// TIA Portal project "000_empty" (V21)

(* hardware
DEVICE "PLC_1"  S7-1500 station
   slot 0: "Rail_0"  Rack  6ES7 590-1***0-0AA0
   slot 1: "PLC_1"  CPU 1513-1 PN  6ES7 513-1AL02-0AB0  V2.9
      slot 3: "CPU display_1"  6ES7591-1AA00-0AA0
      slot 32768: "PROFINET interface_1"  X1
         slot 32769: "Port_1"  X1 P1
         slot 32770: "Port_2"  X1 P2
      slot 34817: "Virtual CP interface port_1"  Virtual CP interface port  Virtual CP interface port
*)

// ===== PLC "PLC_1"  CPU 1513-1 PN =====

TYPE "UDT_Motor"
   STRUCT
      Running : Bool;   // Motor on
      Speed : Real := 1500.0;   // Speed setpoint
      Count : Int := 7;
   END_STRUCT;
END_TYPE

DATA_BLOCK "DB_Global"   // DB1
{ S7_Optimized_Access := 'TRUE' }
   VAR
      xBool : Bool := TRUE;   // Bool comment
      iInt : Int := 42;
      rReal : Real := 3.5;   // Real comment
      aInt : Array[0..3] of Int;
      sData : Struct
         "a" : Bool;
         "b" : DInt := -5;
      END_STRUCT;
   END_VAR
BEGIN
   aInt[1] := 11;
END_DATA_BLOCK

DATA_BLOCK "FB_Empty_DB"   // DB2
{ S7_Optimized_Access := 'TRUE' }
VERSION : 0.1
// stored: InstanceOfName FB_Empty
"FB_Empty"
BEGIN
END_DATA_BLOCK

DATA_BLOCK "DB_Motor"   // DB4
{ S7_Optimized_Access := 'TRUE' }
   VAR
      motor : "UDT_Motor";
   END_VAR
BEGIN
   motor.Speed := 750.0;
END_DATA_BLOCK

// folder: BlockGroup_1

DATA_BLOCK "DB_InGroup"   // DB3
{ S7_Optimized_Access := 'TRUE' }
   VAR
      wWord : Word := 16#00FF;
   END_VAR
BEGIN
END_DATA_BLOCK

// folder: (top level)

FUNCTION_BLOCK "FB_Empty"   // FB1, SCL
{ S7_Optimized_Access := 'TRUE' }
VERSION : 0.1
BEGIN
END_FUNCTION_BLOCK

FUNCTION_BLOCK "FB_Iface"   // FB2, SCL
{ S7_Optimized_Access := 'TRUE' }
VERSION : 0.1
   VAR_INPUT
      iBool : Bool;   // Input bool
      iInt : Int;   // Input int
      iReal : Real;   // Input real
      iArr : Array[0..3] of Int;   // Input array
      iMotor : "UDT_Motor";   // Input UDT
   END_VAR
   VAR_OUTPUT
      oBool : Bool;   // Output bool
      oInt : Int;   // Output int
   END_VAR
   VAR_IN_OUT
      ioReal : Real;   // InOut real
   END_VAR
   VAR
      stInt : Int := 42;   // Static int
      stBool : Bool;   // Static bool comment
   END_VAR
   VAR_TEMP
      tInt : Int;   // Temp int
   END_VAR
   VAR CONSTANT
      cInt : Int := 7;   // Constant int
   END_VAR
BEGIN
   #tInt := #iInt + #cInt;
           #oInt := #tInt;
           #oBool := #iBool;
           #ioReal := #ioReal + #iReal;
END_FUNCTION_BLOCK

FUNCTION "FC_Iface" : Int   // FC1, SCL
{ S7_Optimized_Access := 'TRUE' }
VERSION : 0.1
   VAR_INPUT
      iBool : Bool;   // Input bool
      iInt : Int;   // Input int
      iReal : Real;   // Input real
      iArr : Array[0..3] of Int;   // Input array
      iMotor : "UDT_Motor";   // Input UDT
   END_VAR
   VAR_OUTPUT
      oBool : Bool;   // Output bool
      oInt : Int;   // Output int
   END_VAR
   VAR_IN_OUT
      ioReal : Real;   // InOut real
   END_VAR
   VAR_TEMP
      tInt : Int;   // Temp int
   END_VAR
   VAR CONSTANT
      cInt : Int := 7;   // Constant int
   END_VAR
BEGIN
   #tInt := #iInt + #cInt;
           #oInt := #tInt;
           #oBool := #iBool;
           #ioReal := #ioReal + #iReal;
           #FC_Iface := #tInt;
END_FUNCTION

ORGANIZATION_BLOCK "Main"   // OB1, LAD, ProgramCycle
TITLE = "Main Program Sweep (Cycle)"
{ S7_Optimized_Access := 'TRUE' }
VERSION : 0.1
   VAR_INPUT
      Initial_Call : Bool;   // Initial call of this OB
      Remanence : Bool;   // =True, if remanent data are available
   END_VAR
BEGIN
END_ORGANIZATION_BLOCK